(* IEC 61131-3 sources: programs/VI-54/VI-54_20171205/VI-54_20171205/Stations/PLC_VI54/VI-54_171014/Class/SafetyBaseFSoE (part 5) *)

              LastRequest := _ReadValues;

#ifdef SAFETY_PROTOCOL_ANALYZER_ACTIVATED
  RecordFrame((#StandardRequest)$^DINT, 1);
#endif

              //copy SDO into write-buffer
              ToStdLib.MemCpy(dest := #p_Handle_SDO_Write^.SDOStructure, source := #StandardRequest, size := (sizeof(SDOHeader.StdHeader.CRC) + StandardRequest.SDOHeader.Len));

              //mark SDO data as valid
              p_Handle_SDO_Write^.us_Status := SAFETY_SDO_DATA_VALID;

              if ( pISafety^.udVersion >= 16#1001 ) then
                SAFETY_iPushSafetyTask();
              end_if;

            elsif (UnsafeReadTransNr >= ReadFramesNeeded) then
              // We have finished all read data, go on with the next step
              UnsafeScheduler := UnsafeSchedulerDiagState;
              LastUnsafeUpdate := ops.tAbsolute;
              UnsafeReadTransNr := 0;
            else
              // time until read is not yet over - go on
              UnsafeScheduler := UnsafeSchedulerDiagState;
            end_if;
          else
            UnsafeScheduler := UnsafeSchedulerDiagState;
          end_if;

       (* ***************************************** *)
          UnsafeSchedulerDiagState:
       (* ***************************************** *)
          // get the diag state (on user demand)
          if DiagVars.UserWantsDiagState then

            // get state via SDO communication
            SDORequestBuffer.StdHeader.CRC  := 0;                                                   // CRC is always 0 in Std communication
            SDORequestBuffer.StdHeader.Cmd  := SBF_SDO_COMMAND_GET_STATE;                            // get-state command
            SDORequestBuffer.StdHeader.Typ  := SDO_STD;                                             // standard frame type
            SDORequestBuffer.StdHeader.SeqNr:= StandardSeqNr OR 16#80;                              // sequence number
            SDORequestBuffer.StdHeader.Len  := 4;                                                   // header
            SDORequestBuffer.ud_Address     := 0;
            SDORequestBuffer.us_Length      := 0;

            LastRequest := _DiagState;

#ifdef SAFETY_PROTOCOL_ANALYZER_ACTIVATED
  RecordFrame((#SDORequestBuffer)$^DINT, 1);
#endif

            //copy SDO into write-buffer
            ToStdLib.MemCpy(dest := #p_Handle_SDO_Write^.SDOStructure, source := #SDORequestBuffer, size := (sizeof(SDOHeader.StdHeader.CRC) + SDORequestBuffer.StdHeader.Len));

            //mark SDO data as valid
            p_Handle_SDO_Write^.us_Status := SAFETY_SDO_DATA_VALID;

            if ( pISafety^.udVersion >= 16#1001 ) then
              SAFETY_iPushSafetyTask();
            end_if;
          else
            UnsafeScheduler := UnsafeSchedulerDiagInfo;
          end_if;

       (* ***************************************** *)
          UnsafeSchedulerDiagInfo:
       (* ***************************************** *)

          // get the diag info (on user demand)
          if DiagVars.UserWantsDiagInfo then

            // get state via SDO communication
            StandardRequest.SDOHeader.CRC  := 0;                                                   // CRC is always 0 in Std communication
            StandardRequest.SDOHeader.Cmd  := SBF_SDO_COMMAND_GET_DIAG_INFO;                        // read command
            StandardRequest.SDOHeader.Typ  := SDO_STD;                                             // standard frame type
            StandardRequest.SDOHeader.SeqNr:= StandardSeqNr OR 16#80;                              // sequence number
            StandardRequest.SDOHeader.Len  := 4 + 1;                                               // header + µC-selection
            StandardRequest.aData[0] := DiagVars.ucChoiceDiagInfo;

            LastRequest := _DiagInfo;

#ifdef SAFETY_PROTOCOL_ANALYZER_ACTIVATED
  RecordFrame((#StandardRequest)$^DINT, 1);
#endif

            //copy SDO into write-buffer
            ToStdLib.MemCpy(dest := #p_Handle_SDO_Write^.SDOStructure, source := #StandardRequest, size := (sizeof(SDOHeader.StdHeader.CRC) + StandardRequest.SDOHeader.Len));

            //mark SDO data as valid
            p_Handle_SDO_Write^.us_Status := SAFETY_SDO_DATA_VALID;

            if ( pISafety^.udVersion >= 16#1001 ) then
              SAFETY_iPushSafetyTask();
            end_if;

          else

            if SchedulerStepNo = 6 then
              UnsafeScheduler := UnsafeSchedulerGetDiagVars;

            elsif SchedulerStepNo = 7 then
              UnsafeScheduler := UnsafeSchedulerGetRetryCounter;
            end_if;

          end_if;
       (* ***************************************** *)
          UnsafeSchedulerGetRetryCounter:
       (* ***************************************** *)
          //read out the retry counters every 10seconds
          if (b_DisableSafetyRetryCnt = FALSE)
          & ((ops.tAbsolute - ud_RetryCntTimeMark) > SBF_RETRY_COUNTER_WAIT_TIME)  then

            SDORequestBuffer.StdHeader.CRC  := 0;                                                         // CRC is always 0 in Std communication
            SDORequestBuffer.StdHeader.Cmd  := SBF_SDO_COMMAND_READ;                                       // read command
            SDORequestBuffer.StdHeader.Typ  := SDO_STD;                                                   // standard frame type
            SDORequestBuffer.StdHeader.SeqNr:= StandardSeqNr OR 16#80;                                    // sequence number
            SDORequestBuffer.StdHeader.Len  := 4 + 4 + SBF_SDO_LENGTH_RETRY_COUNTER;                       // header + destination address + length of data
            SDORequestBuffer.ud_Address     := SBF_SDO_ADDRESS_RETRY_COUNTER;                              // address of retrycounter
            SDORequestBuffer.us_Length      := SBF_SDO_LENGTH_RETRY_COUNTER;                               // length of data

            LastRequest := _ReadRetryCounter;

  #ifdef SAFETY_PROTOCOL_ANALYZER_ACTIVATED
  RecordFrame((#SDORequestBuffer)$^DINT, 1);
  #endif

            //copy SDO into write-buffer
            ToStdLib.MemCpy(dest := #p_Handle_SDO_Write^.SDOStructure, source := #SDORequestBuffer, size := (sizeof(SDOHeader.StdHeader.CRC) + SDORequestBuffer.StdHeader.Len));

            //mark SDO data as valid
            p_Handle_SDO_Write^.us_Status := SAFETY_SDO_DATA_VALID;

            if ( pISafety^.udVersion >= 16#1001 ) then
              SAFETY_iPushSafetyTask();
            end_if;

            //reset timemark
            ud_RetryCntTimeMark := ops.tAbsolute;

          else
            UnsafeScheduler := UnsafeSchedulerGetDiagVars;
          end_if;
        else
          LogError("Undefined Scheduler-State");
        end_case;
      end_while;
    end_if;
  end_if;

  // at the first run we write all variables independent of any changes
  if RunState > OldRunState then
    SendAllUnsafeValues();
  end_if;
  OldRunState := RunState;

	state := READY;

//============================ Profiler start======================================================
#ifdef  DM_Profiler
  StopTimeMeasurement(usMode := DMTIME_CY);
#endif
//============================ Profiler end========================================================
END_FUNCTION

FUNCTION VIRTUAL SafetyBaseFSoE::GetConfiguration

END_FUNCTION

FUNCTION VIRTUAL SafetyBaseFSoE::SetSafetyState
	VAR_INPUT
		NewState 	: SafetyConfigStateType;
	END_VAR

  // use it locally => can also be forwarded in derivation
  SafetyState := NewState;

END_FUNCTION

FUNCTION VIRTUAL SafetyBaseFSoE::RefreshAsySrv
  // derive this
END_FUNCTION

FUNCTION VIRTUAL SafetyBaseFSoE::SetRetryCounter

  SafetyRetryCounter := -1;

END_FUNCTION

FUNCTION SafetyBaseFSoE::IsInCache
	VAR_INPUT
		ud_Address 	: UDINT;
		us_Length 	: USINT;
	END_VAR
	VAR_OUTPUT
		ItsInside 	: BOOL;
	END_VAR

  if CachedSize &
     (ud_Address >= CachedAddr) &
     ((ud_Address + us_Length) <= (CachedAddr + CachedSize)) then
    ItsInside := TRUE;
  else
    ItsInside := FALSE;
  end_if;

END_FUNCTION

FUNCTION SafetyBaseFSoE::AddToCache
	VAR_INPUT
		p_SDORequestBuffer 	: ^SDORequReadConfig;
		p_SDOResponseBuffer 	: ^SDORespReadConfig;
	END_VAR

  if p_SDORequestBuffer^.us_Length then
    CachedAddr := p_SDORequestBuffer^.ud_Address;
    CachedSize := p_SDORequestBuffer^.us_Length;
    _memcpy(ptr1:=#Cache, ptr2:=#p_SDOResponseBuffer^.ud_Data, cntr:=p_SDORequestBuffer^.us_Length);
  end_if;

END_FUNCTION

FUNCTION SafetyBaseFSoE::GetFSoEConnectionInfos
	VAR_INPUT
		p_SDORequestBuffer 	: ^SafetyBaseFSoE::SDORequReadConfig;
		p_SDOResponseBuffer 	: ^SafetyBaseFSoE::SDORespReadConfig;
	END_VAR
  VAR
  	Address         : UDINT;
    Size            : USINT;
    sd_retval       : DINT;
    i               : UDINT;
    pActConnection  : ^t_FSoEConnectionDetails;
    TempRoutingInfo : t_FSoERoutingInfoElement;
    NextAddress     : UDINT;
  END_VAR

  // free the list if there is still one
  FreeFSoEConnectionInfos();

  // check if we already got the info:
  if ConnectionInfos.ConnectionNo | ConnectionInfos.pFirstConnection then
    LogError("(SafetyBaseFSoE::GetFSoEConnectionInfos) List already exists! May not have been resetted correctly!");
    return;
  end_if;

//*****************************************************************************
//** CONNECTION STATE INFO                                                   **
//*****************************************************************************

  // get number of connections
  Address := SBF_SDO_ADDRESS_FSOE_CONN_STATE;
  Size    := 2;

  //send request and receive data
  sd_retval := SDOReadCfgRequ ( p_SDORequestBuffer  := p_SDORequestBuffer
                              , p_SDOResponseBuffer := p_SDOResponseBuffer
                              , ud_Address          := Address
                              , us_Length           := Size
                              );

  //no response
  if ( sd_retval <> 0 ) then
    LogError("(SafetyBaseFSoE::GetFSoEConnectionInfos) Config Read Error: Error reading number of connections");
    return;
  end_if;

  ConnectionInfos.ConnectionNo := p_SDOResponseBuffer^.ud_Data$UINT;

  if ConnectionInfos.ConnectionNo = 0 then
    // no connections available
    return;
  end_if;

  // allocate memory for the connections
  ConnectionInfos.pFirstConnection$pVoid := ToStdLib.Malloc(size:= ConnectionInfos.ConnectionNo * sizeof(t_FSoEConnectionDetails));

  if ConnectionInfos.pFirstConnection = NIL then
    LogError("(SafetyBaseFSoE::GetFSoEConnectionInfos) Config Read Error: Failed to allocate memory for FSoE connection details");
    return;
  end_if;

  // reset memory (also resets pNext although we are not using a linked list here)
  _memset(dest:=ConnectionInfos.pFirstConnection, usByte:=0, cntr:= ConnectionInfos.ConnectionNo * sizeof(t_FSoEConnectionDetails));

  Address += Size;
  Size    := 1;

  pActConnection := ConnectionInfos.pFirstConnection;

  // get connection states
  for i := 0 to ConnectionInfos.ConnectionNo-1 do
    // get state of connection

    //send request and receive data
    sd_retval := SDOReadCfgRequ ( p_SDORequestBuffer  := p_SDORequestBuffer
                                , p_SDOResponseBuffer := p_SDOResponseBuffer
                                , ud_Address          := Address
                                , us_Length           := Size
                                );

    //no response
    if ( sd_retval <> 0 ) then
      LogError("(SafetyBaseFSoE::GetFSoEConnectionInfos) Config Read Error: Error reading connection state");
      return;
    end_if;

    // get connection state
    pActConnection^.ConnectionState := (p_SDOResponseBuffer^.ud_Data$USINT AND 2#0111)$t_FSoEConnectionState;

    // get info if the module is master or slave at this connection
    pActConnection^.Flags.IsMaster  := (p_SDOResponseBuffer^.ud_Data$USINT AND 2#1000) <> 0;

    // save safety number
    pActConnection^.OwnerSafetyNbr  := SafetyNumber;

    // for easier debugging we set the correct next pointers
    if i = ConnectionInfos.ConnectionNo-1 then
      pActConnection^.pNext := NIL;
    else
      pActConnection^.pNext := pActConnection + sizeof(t_FSoEConnectionDetails);
    end_if;

    pActConnection                  += sizeof(t_FSoEConnectionDetails);
    Address                         += Size;
  end_for;

//*****************************************************************************
//** ROUTING INFO                                                            **
//*****************************************************************************

  // get number of connections
  Address := SBF_SDO_ADDRESS_FSOE_ROUTING_INFO;
  Size    := 2;

  //send request and receive data
  sd_retval := SDOReadCfgRequ ( p_SDORequestBuffer  := p_SDORequestBuffer
                              , p_SDOResponseBuffer := p_SDOResponseBuffer
                              , ud_Address          := Address
                              , us_Length           := Size
                              );

  //no response
  if ( sd_retval <> 0 ) then
    LogError("(SafetyBaseFSoE::GetFSoEConnectionInfos) Config Read Error: Error reading number of connections");
    return;
  end_if;

  // check if it's the same number
  if ConnectionInfos.ConnectionNo <> p_SDOResponseBuffer^.ud_Data$UINT then
    LogError("(SafetyBaseFSoE::GetFSoEConnectionInfos) Config Read Error: Number of connections does not match (case 1)");
    return;
  end_if;

  Address += Size;
  Size    := sizeof(t_FSoERoutingInfoElement);

  pActConnection := ConnectionInfos.pFirstConnection;

  // get connection states
  for i := 0 to ConnectionInfos.ConnectionNo-1 do
    // get routing info of connections

    //send request and receive data
    sd_retval := SDOReadCfgRequ ( p_SDORequestBuffer  := p_SDORequestBuffer
                                , p_SDOResponseBuffer := p_SDOResponseBuffer
                                , ud_Address          := Address
                                , us_Length           := Size
                                );

    //no response
    if ( sd_retval <> 0 ) then
      LogError("(SafetyBaseFSoE::GetFSoEConnectionInfos) Config Read Error: Error reading routing info");
      return;
    end_if;

    TempRoutingInfo := p_SDOResponseBuffer^.ud_Data$t_FSoERoutingInfoElement;

    // store the data in the connection info
    pActConnection^.SlaveAddress        := TempRoutingInfo.SlaveAddress;
    pActConnection^.MasterReadSize      := TempRoutingInfo.SafeOutputFrameSize;
    pActConnection^.MasterWriteSize     := TempRoutingInfo.SafeInputFrameSize;

    // the offset info depends on if we are master or slave
    if pActConnection^.Flags.IsMaster then
      pActConnection^.MasterReadOffset  := TempRoutingInfo.SafeOutputFrameOffset;
      pActConnection^.MasterWriteOffset := TempRoutingInfo.SafeInputFrameOffset;
    else
      pActConnection^.SlaveWriteOffset  := TempRoutingInfo.SafeOutputFrameOffset;
      pActConnection^.SlaveReadOffset   := TempRoutingInfo.SafeInputFrameOffset;
    end_if;

    pActConnection                  += sizeof(t_FSoEConnectionDetails);
    Address                         += Size;
  end_for;

//*****************************************************************************
//** CONNECTION INSTANCES                                                    **
//*****************************************************************************

  Address := SBF_SDO_ADDRESS_FSOE_CONN_INST;
  Size    := 4;

  //send request and receive data
  sd_retval := SDOReadCfgRequ ( p_SDORequestBuffer  := p_SDORequestBuffer
                              , p_SDOResponseBuffer := p_SDOResponseBuffer
                              , ud_Address          := Address
                              , us_Length           := Size
                              );

  //no response
  if ( sd_retval <> 0 ) then
    LogError("(SafetyBaseFSoE::GetFSoEConnectionInfos) Config Read Error: Error reading number of connections");
    return;
  end_if;

  // check if it's the same number
  if ConnectionInfos.ConnectionNo <> p_SDOResponseBuffer^.ud_Data then
    LogError("(SafetyBaseFSoE::GetFSoEConnectionInfos) Config Read Error: Number of connections does not match (case 2)");
    return;
  end_if;

  Address += Size;

  pActConnection := ConnectionInfos.pFirstConnection;

  // get connection states
  for i := 0 to ConnectionInfos.ConnectionNo-1 do
    // get routing instance info of connections

    Size := 4;

    //send request and receive data
    sd_retval := SDOReadCfgRequ ( p_SDORequestBuffer  := p_SDORequestBuffer
                                , p_SDOResponseBuffer := p_SDOResponseBuffer
                                , ud_Address          := Address
                                , us_Length           := Size
                                );

    //no response
    if ( sd_retval <> 0 ) then
      LogError("(SafetyBaseFSoE::GetFSoEConnectionInfos) Config Read Error: Error reading size of routing instance info");
      return;
    end_if;

    // calculate address of next connection (to check it later)
    NextAddress := Address + p_SDOResponseBuffer^.ud_Data;

    // get the flags
    Address   += Size;
    Size      := 4;

    //send request and receive data
    sd_retval := SDOReadCfgRequ ( p_SDORequestBuffer  := p_SDORequestBuffer
                                , p_SDOResponseBuffer := p_SDOResponseBuffer
                                , ud_Address          := Address
                                , us_Length           := Size
                                );

    //no response
    if ( sd_retval <> 0 ) then
      LogError("(SafetyBaseFSoE::GetFSoEConnectionInfos) Config Read Error: Error reading flags of routing instance info");
      return;
    end_if;

    if ((p_SDOResponseBuffer^.ud_Data AND 1) <> 0) <> pActConnection^.Flags.IsMaster then
      LogError("(SafetyBaseFSoE::GetFSoEConnectionInfos) Config Read Error: Master settings mismatch");
      return;
    end_if;

    pActConnection^.Flags := p_SDOResponseBuffer^.ud_Data$USINT;

    // get the net size of the safe output data (only the bits for the I/Os without crc and stuff)
    Address   += Size;
    Size      := 2;

    //send request and receive data
    sd_retval := SDOReadCfgRequ ( p_SDORequestBuffer  := p_SDORequestBuffer
                                , p_SDOResponseBuffer := p_SDOResponseBuffer
                                , ud_Address          := Address
                                , us_Length           := Size
                                );

    //no response
    if ( sd_retval <> 0 ) then
      LogError("(SafetyBaseFSoE::GetFSoEConnectionInfos) Config Read Error: Error reading safe output net size of routing instance info");
      return;
    end_if;

    // we don't need the net size yet

    // get the net size of the safe input data (only the bits for the I/Os without crc and stuff)
    Address   += Size;
    Size      := 2;

    //send request and receive data
    sd_retval := SDOReadCfgRequ ( p_SDORequestBuffer  := p_SDORequestBuffer
                                , p_SDOResponseBuffer := p_SDOResponseBuffer
                                , ud_Address          := Address
                                , us_Length           := Size
                                );

    //no response
    if ( sd_retval <> 0 ) then
      LogError("(SafetyBaseFSoE::GetFSoEConnectionInfos) Config Read Error: Error reading safe input net size of routing instance info");
      return;
    end_if;

    // we don't need the net size yet

    // get the slave address
    Address   += Size;
    Size      := 2;

    //send request and receive data
    sd_retval := SDOReadCfgRequ ( p_SDORequestBuffer  := p_SDORequestBuffer
                                , p_SDOResponseBuffer := p_SDOResponseBuffer
                                , ud_Address          := Address
                                , us_Length           := Size
                                );

    //no response
    if ( sd_retval <> 0 ) then
      LogError("(SafetyBaseFSoE::GetFSoEConnectionInfos) Config Read Error: Error reading slave address of routing instance info");
      return;
    end_if;

    // the following settings are only available in the master
    if pActConnection^.Flags.IsMaster then

      // get the connection ID
      Address   += Size;
      Size      := 2;

      //send request and receive data
      sd_retval := SDOReadCfgRequ ( p_SDORequestBuffer  := p_SDORequestBuffer
                                  , p_SDOResponseBuffer := p_SDOResponseBuffer
                                  , ud_Address          := Address
                                  , us_Length           := Size
                                  );

      //no response
      if ( sd_retval <> 0 ) then
        LogError("(SafetyBaseFSoE::GetFSoEConnectionInfos) Config Read Error: Error reading the connection ID of routing instance info");
        return;
      end_if;

      pActConnection^.ConnectionID := p_SDOResponseBuffer^.ud_Data$UINT;

      // get transmission time
      Address   += Size;
      Size      := 2;

      //send request and receive data
      sd_retval := SDOReadCfgRequ ( p_SDORequestBuffer  := p_SDORequestBuffer
                                  , p_SDOResponseBuffer := p_SDOResponseBuffer
                                  , ud_Address          := Address
                                  , us_Length           := Size
                                  );

      //no response
      if ( sd_retval <> 0 ) then
        LogError("(SafetyBaseFSoE::GetFSoEConnectionInfos) Config Read Error: Error reading the transmission time of routing instance info");
        return;
      end_if;

      pActConnection^.TransmissionTime_ms := p_SDOResponseBuffer^.ud_Data$UINT;

      // get length of communication parameters (must be 2)
      Address   += Size;
      Size      := 2;

      //send request and receive data
      sd_retval := SDOReadCfgRequ ( p_SDORequestBuffer  := p_SDORequestBuffer
                                  , p_SDOResponseBuffer := p_SDOResponseBuffer
                                  , ud_Address          := Address
                                  , us_Length           := Size
                                  );

      //no response
      if ( sd_retval <> 0 ) then
        LogError("(SafetyBaseFSoE::GetFSoEConnectionInfos) Config Read Error: Error reading the length of the communication parameters of routing instance info");
        return;
      end_if;

      if p_SDOResponseBuffer^.ud_Data$UINT <> 2 then
        LogError("(SafetyBaseFSoE::GetFSoEConnectionInfos) Config Read Error: Length of communication parameters is wrong");
        return;
      end_if;

      // skip FSoE watchdog time in ms
      Address   += Size;
      Size      := 2;

      // get size of application parameters
      Address   += Size;
      Size      := 2;

      //send request and receive data
      sd_retval := SDOReadCfgRequ ( p_SDORequestBuffer  := p_SDORequestBuffer
                                  , p_SDOResponseBuffer := p_SDOResponseBuffer
                                  , ud_Address          := Address
                                  , us_Length           := Size
                                  );

      //no response
      if ( sd_retval <> 0 ) then
        LogError("(SafetyBaseFSoE::GetFSoEConnectionInfos) Config Read Error: Error reading the length of the application parameters of routing instance info");
        return;
      end_if;

      // skip length
      Address   += Size;

      // skip application parameters
      Size      := p_SDOResponseBuffer^.ud_Data$USINT;
      Address   += Size;

      // get to a 4 byte aligned address
      if (Address MOD 4) then
        Address := Address + (4 - (Address MOD 4)); //increase memory, up to a value, which could be divided by 4
      end_if;

      // get size of hw path
      Size      := 4;

      //send request and receive data
      sd_retval := SDOReadCfgRequ ( p_SDORequestBuffer  := p_SDORequestBuffer
                                  , p_SDOResponseBuffer := p_SDOResponseBuffer
                                  , ud_Address          := Address
                                  , us_Length           := Size
                                  );

      //no response
      if ( sd_retval <> 0 ) then
        LogError("(SafetyBaseFSoE::GetFSoEConnectionInfos) Config Read Error: Error reading the hardware path length of routing instance info");
        return;
      end_if;

      // get the hardware path
      Address   += Size;
      Size      := p_SDOResponseBuffer^.ud_Data$USINT;

      if Size = 0 then
        LogError("(SafetyBaseFSoE::GetFSoEConnectionInfos) Config Read Error: Hardware path length is zero");
        return;
      end_if;

      //send request and receive data
      sd_retval := SDOReadCfgRequ ( p_SDORequestBuffer  := p_SDORequestBuffer
                                  , p_SDOResponseBuffer := p_SDOResponseBuffer
                                  , ud_Address          := Address
                                  , us_Length           := Size
                                  );

      //no response
      if ( sd_retval <> 0 ) then
        LogError("(SafetyBaseFSoE::GetFSoEConnectionInfos) Config Read Error: Error reading the hardware path of routing instance info");
        return;
      end_if;

      // save hardware path into structure
      pActConnection^.SlavePathLen      := Size;
      pActConnection^.pSlavePath$pVoid  := ToStdLib.Malloc(size:=Size);

      if pActConnection^.pSlavePath = NIL then
        LogError("(SafetyBaseFSoE::GetFSoEConnectionInfos) Failed to allocate memory for the slave hardware path at the routing instance info");
        return;
      end_if;

      _memcpy(ptr1:=pActConnection^.pSlavePath, ptr2:=#p_SDOResponseBuffer^.ud_Data, cntr:=pActConnection^.SlavePathLen);

      Address         += Size;

      // get to a 4 byte aligned address
      if (Address MOD 4) then
        Address := Address + (4 - (Address MOD 4)); //increase memory, up to a value, which could be divided by 4
      end_if;

      // get size of compressed hw path
      Size      := 4;

      //send request and receive data
      sd_retval := SDOReadCfgRequ ( p_SDORequestBuffer  := p_SDORequestBuffer
                                  , p_SDOResponseBuffer := p_SDOResponseBuffer
                                  , ud_Address          := Address
                                  , us_Length           := Size
                                  );

      //no response
      if ( sd_retval <> 0 ) then
        LogError("(SafetyBaseFSoE::GetFSoEConnectionInfos) Config Read Error: Error reading the compressed hardware path length of routing instance info");
        return;
      end_if;

      // get the hardware path
      Address   += Size;
      Size      := p_SDOResponseBuffer^.ud_Data$USINT;

      //send request and receive data
      sd_retval := SDOReadCfgRequ ( p_SDORequestBuffer  := p_SDORequestBuffer
                                  , p_SDOResponseBuffer := p_SDOResponseBuffer
                                  , ud_Address          := Address
                                  , us_Length           := Size
                                  );

      //no response
      if ( sd_retval <> 0 ) then
        LogError("(SafetyBaseFSoE::GetFSoEConnectionInfos) Config Read Error: Error reading the compressed hardware path of routing instance info");
        return;
      end_if;

      // save compressed hardware path into structure
      pActConnection^.SlavePathCompLen      := Size;
      pActConnection^.pSlavePathComp$pVoid  := ToStdLib.Malloc(size:=Size);

      if pActConnection^.pSlavePathComp = NIL then
        LogError("(SafetyBaseFSoE::GetFSoEConnectionInfos) Failed to allocate memory for the compressed slave hardware path at the routing instance info");
        return;
      end_if;

      _memcpy(ptr1:=pActConnection^.pSlavePathComp, ptr2:=#p_SDOResponseBuffer^.ud_Data, cntr:=pActConnection^.SlavePathCompLen);

      Address         += Size;

      // get to a 4 byte aligned address
      if (Address MOD 4) then
        Address := Address + (4 - (Address MOD 4)); //increase memory, up to a value, which could be divided by 4
      end_if;

      if Address > NextAddress then
        LogError("(SafetyBaseFSoE::GetFSoEConnectionInfos) Config Read Error: Structure size mismatch");
        return;
      end_if;
    end_if;

    Address         := NextAddress;
    pActConnection  += sizeof(t_FSoEConnectionDetails);
  end_for;

END_FUNCTION

FUNCTION SafetyBaseFSoE::FreeFSoEConnectionInfos
  VAR
    i               : UDINT;
    pActConnection  : ^t_FSoEConnectionDetails;
  END_VAR

  if (ConnectionInfos.ConnectionNo = 0) | (ConnectionInfos.pFirstConnection = NIL) then
    // nothing to free
    return;
  end_if;

  // check if all connections have been initialized
  pActConnection := ConnectionInfos.pFirstConnection;
  for i := 0 to ConnectionInfos.ConnectionNo-1 do
    if pActConnection^.ConnectionState = FCS_NOT_INITIALIZED then
      // not yet time to free them
      return;
    end_if;

    pActConnection += sizeof(t_FSoEConnectionDetails);
  end_for;

  pActConnection := ConnectionInfos.pFirstConnection;
  for i := 0 to ConnectionInfos.ConnectionNo-1 do
    // free hardware path memory

    if pActConnection^.pSlavePath then
      ToStdLib.Free(mptr:=pActConnection^.pSlavePath);
    end_if;

    if pActConnection^.pSlavePathComp then
      ToStdLib.Free(mptr:=pActConnection^.pSlavePathComp);
    end_if;

    pActConnection += sizeof(t_FSoEConnectionDetails);
  end_for;

  // free the connectionlist
  ToStdLib.Free(mptr:=ConnectionInfos.pFirstConnection);
  ConnectionInfos.pFirstConnection := NIL;
  ConnectionInfos.ConnectionNo := 0;

END_FUNCTION

FUNCTION SafetyBaseFSoE::CheckFSoEConnections
  VAR
		MyPara 	            : CmdStruct;
		MyResult	          : results;
    i                   : UDINT;
    pActConnection      : ^t_FSoEConnectionDetails;
    SDORequestBuffer    : SDORequReadConfig;
    SDOResponseBuffer   : ARRAY [0..SBF_SDO_MAX_LENGTH-1] OF USINT;
		p_SDORequestBuffer 	: ^SDORequReadConfig;
		p_SDOResponseBuffer : ^SDORespReadConfig;
    UnInifializedNo     : UDINT;
    sd_retval           : DINT;
  END_VAR

  // there were some of the FSoE connections not initialized when fetching the configuration data => update them

  UnInifializedNo := 0;

  //SDO request for this command has 5 bytes additional to the header
  p_SDORequestBuffer := #SDORequestBuffer;

  //SDO response for this command can have maximum additional data
  p_SDOResponseBuffer := (#SDOResponseBuffer)$^SDORespReadConfig;

  //calculate length without crc
  p_SDORequestBuffer^.StdHeader.Len := sizeof(SDORequReadConfig) - sizeof(SDOHeader.StdHeader.CRC);

  //type
  p_SDORequestBuffer^.StdHeader.Typ := SDO_STD;

  //command for reading config data
  p_SDORequestBuffer^.StdHeader.Cmd := SBF_SDO_COMMAND_READ;

  // reset cache, because it may contain an old access on the same address => we want fresh data
  CachedSize := 0;

  pActConnection := ConnectionInfos.pFirstConnection;

  for i := 0 to ConnectionInfos.ConnectionNo-1 do
    if pActConnection^.ConnectionState = FCS_NOT_INITIALIZED then
      UnInifializedNo += 1;

      //send request and receive data
      sd_retval := SDOReadCfgRequ ( p_SDORequestBuffer  := p_SDORequestBuffer
                                  , p_SDOResponseBuffer := p_SDOResponseBuffer
                                  , ud_Address          := SBF_SDO_ADDRESS_FSOE_CONN_STATE + 2 + i
                                  , us_Length           := 1
                                  );

      //no response
      if ( sd_retval <> 0 ) then
        LogError("(SafetyBaseFSoE::CheckFSoEConnections) Config Read Error: Error reading connection state");
        return;
      end_if;

      // get connection state
      pActConnection^.ConnectionState := (p_SDOResponseBuffer^.ud_Data$USINT AND 2#0111)$t_FSoEConnectionState;

      if pActConnection^.ConnectionState <> FCS_NOT_INITIALIZED then
        UnInifializedNo -= 1;

        // get the corresponding slave address number

        //send request and receive data
        sd_retval := SDOReadCfgRequ ( p_SDORequestBuffer  := p_SDORequestBuffer
                                    , p_SDOResponseBuffer := p_SDOResponseBuffer
                                    , ud_Address          := SBF_SDO_ADDRESS_FSOE_ROUTING_INFO + 2 + i * sizeof(t_FSoERoutingInfoElement)
                                    , us_Length           := sizeof(t_FSoERoutingInfoElement)
                                    );

        //no response
        if ( sd_retval <> 0 ) then
          LogError("(SafetyBaseFSoE::CheckFSoEConnections) Config Read Error: Error reading routing info");
          return;
        end_if;

        pActConnection^.SlaveAddress := p_SDOResponseBuffer^.ud_Data$t_FSoERoutingInfoElement.SlaveAddress;

        if pActConnection^.SlaveAddress = 0 then
          LogError(e_msg:="(SafetyBaseFSoE::CheckFSoEConnections) Connection initialized but slave address is still zero!");
        end_if;
      end_if;
    end_if;

    pActConnection                  += sizeof(t_FSoEConnectionDetails);
  end_for;

  // if all connections are initialized => tell the safety manager
  if (UnInifializedNo = 0) & pSafetyManagerThis then
    MyPara.uiCmd    := CMD_SM_FSOE_CON_INITIALIZED;
    MyPara.aPara[0] := SafetyNumber$DINT;
    MyPara.aPara[1] := ConnectionInfos.ConnectionNo$DINT;
    MyPara.aPara[2] := ConnectionInfos.pFirstConnection$DINT;

    if pSafetyManagerThis^.NewInst(#MyPara, #MyResult) = READY then
      // we don't need this memory anymore
      FreeFSoEConnectionInfos();
    end_if;
  end_if;

END_FUNCTION

FUNCTION VIRTUAL GLOBAL SafetyBaseFSoE::GetDiagConnect::NewInst
	VAR_INPUT
		pPara 	: ^CmdStruct;
		pResult 	: ^Results;
	END_VAR
	VAR_OUTPUT
		ret_code 	: IprStates;
	END_VAR

	ret_code := READY;

	CASE pPara^.uiCmd OF

    CMD_SM_DIAG_GET_INFO:

      //Subcommand
      case pPara^.aPara[0] of
//*****************************************************************************
        SBCMD_SM_DIAG_GET_INFO:
          pResult^.aData[0] :=  GetDiagInfo(pDiagInfo:=(pPara^.aPara[1])$^SafetyDiagInfo);

//*****************************************************************************
        SBCMD_SM_DIAG_GET_STATE:
          pResult^.aData[0] :=  GetDiagState(pDiagState:=(pPara^.aPara[1])$^SafetyDiagState);

//*****************************************************************************
        SBCMD_SM_DIAG_FETCH_INFO:
      //Fetch Diag Info for uCx
          FetchDiagInfo(ucChoice:=pPara^.aPara[1]$USINT);

//*****************************************************************************
        SBCMD_SM_DIAG_FETCH_STATE:
      FetchDiagState();

//*****************************************************************************
        SBCMD_SM_DIAG_IS_SAVE_LOG_ACTIVE:
      pResult^.aData[0] := SaveLogActive();

//*****************************************************************************
        SBCMD_SM_DIAG_SAVE_LOGFILE:
          pResult^.aData[0] := (SaveLog(ucChoice:=(pPara^.aPara[1])$USINT, pDPNE:=(pPara^.aPara[2])$^CHAR))$USINT;

//*****************************************************************************
        SBCMD_SM_DIAG_GET_SAVE_LOGFILE_STATE:
      pResult^.aData[0] := DiagVars.SavingLogSuccessful$USINT;

//*****************************************************************************
        SBCMD_SM_DIAG_GET_SAFETY_NUMBER:
      pResult^.aData[0]$UDINT := SafetyNumber;

//*****************************************************************************
        SBCMD_SM_DIAG_GET_SAFETY_STATE:
      pResult^.aData[0] := SafetyState$USINT;

//*****************************************************************************
        SBCMD_SM_DIAG_IS_DIAGNOSE_AVAILABLE:
          pResult^.aData[0] := TRUE;

	END_CASE;
    else
      TRACE("(SafetyBaseFSoE::GetDiagConnect::NewInst) Unknown command!");
      ret_code := ERROR;
	END_CASE;

END_FUNCTION

FUNCTION SafetyBaseFSoE::GetNewMemSize
	VAR_INPUT
		Required 	: UDINT;
	END_VAR
	VAR_OUTPUT
		NextBiggerBlockSize 	: UDINT;
	END_VAR

  // how many complete blocks are necessary
  NextBiggerBlockSize := Required / SBF_CONFIG_MEMORY_BLOCK_SIZE;

  // is there also an incomplete block?
  if Required MOD SBF_CONFIG_MEMORY_BLOCK_SIZE then
    NextBiggerBlockSize += 1;
  end_if;

  // now that we have the number of blocks necessary => get number of bytes
  NextBiggerBlockSize *= SBF_CONFIG_MEMORY_BLOCK_SIZE;

END_FUNCTION

FUNCTION SafetyBaseFSoE::CheckAddDynSlaveResponse
	VAR_INPUT
		pAddDynSlaveRsp 	: ^t_AddDynSlaveResponse;
	END_VAR
	VAR_OUTPUT
		ResponseOk 	: BOOL;
	END_VAR

  // check if any of the offset/length combination exceeds our access to the module
  if ((pAddDynSlaveRsp^.OffsetSafeInData  + pAddDynSlaveRsp^.LenSafeInData ) > MyPDOWriteSize) |
     ((pAddDynSlaveRsp^.OffsetSafeOutData + pAddDynSlaveRsp^.LenSafeOutData) > MyPDOReadSize ) then
    ResponseOk := FALSE;

    LogError("CheckAddDynSlaveResponse: Invalid offset/length combination of read or write data in AddDynSlave response");
  else
    ResponseOk := TRUE;
  end_if;

END_FUNCTION
